// TIA Portal V21 export
// export: Created 2026-10-23T20:42:47.6019008Z, ExportSetting WithDefaults, DisplayName Totally Integrated Automation Portal, DisplayVersion V21 Update 1, DisplayName SINAMICS Startdrive Advanced, DisplayVersion V21 HF2, DisplayName SINAMICS Startdrive G110M, G120, G120C, G120D, G120P, G115D, DisplayVersion V21 HF2, DisplayName SINAMICS Startdrive G130, G150, S120, S150, G200, G220, S200, S210, S220, Innomotics MVD, DisplayVersion V21 HF2, DisplayName STEP 7 Professional, DisplayVersion V21 Update 1, DisplayName STEP 7 Safety, DisplayVersion V21, DisplayName Tech WebApplication, DisplayVersion V21, DisplayName WinCC Basic/Comfort/Advanced, DisplayVersion V21 Update 1, DisplayName WinCC Unified, DisplayVersion V21 Update 1
FUNCTION_BLOCK "FB_FbdBoxes"   // FB10, FBD
TITLE = FUP-Boxen, Aufruf und Sprung / FBD boxes, call and jump
{ S7_Optimized_Access := 'TRUE' }
VERSION : 0.1
// TON, MOVE, ADD, Vergleich, FB-Aufruf mit EN/ENO und ein Sprung mit Marke in FUP / TON, MOVE, ADD, compare, FB call with EN/ENO and a jump with label in FBD
// stored: AutoNumber true, IsIECCheckEnabled false, IsRetainMemResEnabled false, MemoryReserve 100, SetENOAutomatically false, UDAEnableTagReadback false
   VAR_INPUT
      Start : Bool;   // Startbefehl / Start command
      InValue : Int;   // Eingangswert / Input value
      Limit : Int := 100;   // Grenzwert für den Vergleich / Limit for the comparison
   END_VAR
   VAR_OUTPUT
      Delayed : Bool;   // Start um drei Sekunden verzögert / Start delayed by three seconds
      Copy : Int;   // Kopie des Eingangswerts / Copy of the input value
      Sum : Int;   // Eingangswert plus Grenzwert / Input value plus limit
      IsEqual : Bool;   // Eingangswert gleich dem Grenzwert / Input value equal to the limit
      SectionsOk : Bool;   // ENO des Aufrufs von FB_SclTimers / ENO of the FB_SclTimers call
      Skipped : Bool;   // Nur gesetzt, wenn nicht gesprungen wird / Set only when the jump is not taken
      AfterJump : Bool;   // Netzwerk nach der Sprungmarke / Network after the jump label
   END_VAR
   VAR
      Delay { S7_SetPoint := 'True'} : TON_TIME;   // Einschaltverzögerung / On-delay timer
      DelayElapsed : Time;   // Abgelaufene Zeit der Einschaltverzögerung / Elapsed time of the on-delay timer
      Timers { S7_SetPoint := 'True'} : "FB_SclTimers";   // Multiinstanz von FB_SclTimers / Multi-instance of FB_SclTimers
      TimerRunOn : Bool;   // Nachlaufausgang von FB_SclTimers / Run-on output of FB_SclTimers
      TimerPulse : Bool;   // Impulsausgang von FB_SclTimers / Pulse output of FB_SclTimers
      TimerCount : Int;   // Zählausgang von FB_SclTimers / Count output of FB_SclTimers
      TimerDelayed : Bool;   // Verzögerter Ausgang von FB_SclTimers / Delayed output of FB_SclTimers
      TimerReached : Bool;   // Ausgang Zählwert erreicht von FB_SclTimers / Count reached output of FB_SclTimers
   END_VAR
   VAR_TEMP   // added for the SCL form of the ladder/FBD networks
      _w1 : Bool;
   END_VAR
BEGIN

REGION Network 1: Einschaltverzögerung als Multiinstanz / On-delay timer as multi-instance
   // Der Ausgang folgt dem Startbefehl nach drei Sekunden. / The output follows the start command after three seconds.
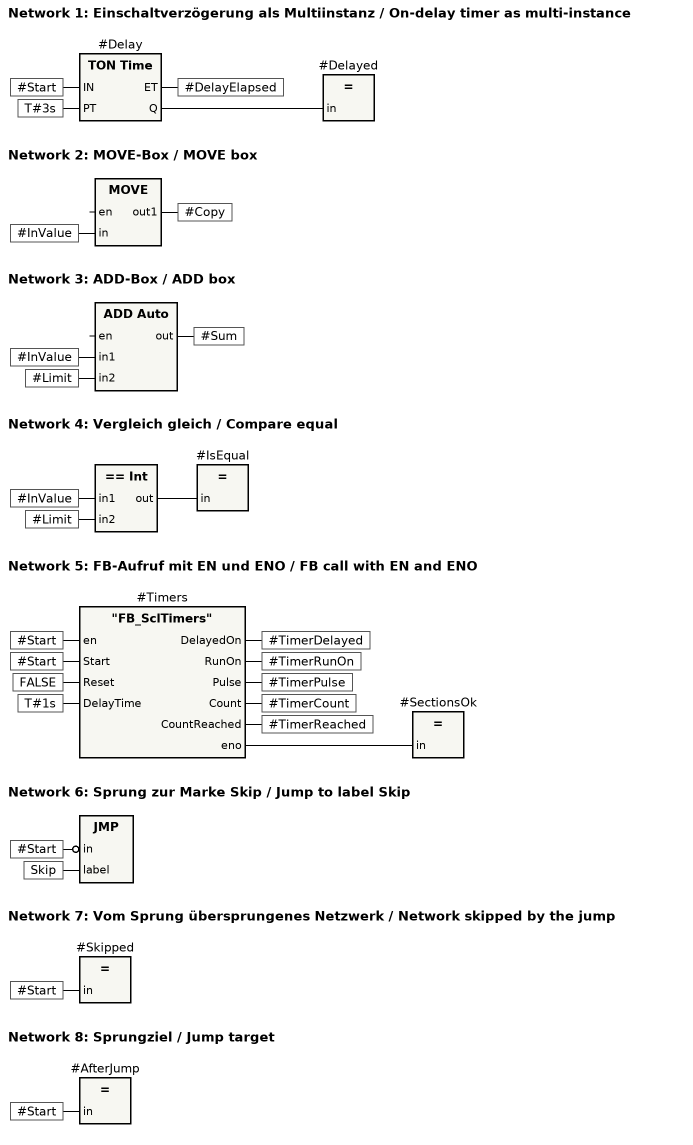
   #Delay(IN := #Start, PT := T#3s, ET => #DelayElapsed);   // TON
   #Delayed := #Delay.Q;
END_REGION

REGION Network 2: MOVE-Box / MOVE box
   // Kopiert den Eingangswert. / Copies the input value.
   #Copy := #InValue;
END_REGION

REGION Network 3: ADD-Box / ADD box
   // Addiert den Grenzwert zum Eingangswert. / Adds the limit to the input value.
   #Sum := #InValue + #Limit;
END_REGION

REGION Network 4: Vergleich gleich / Compare equal
   // Wahr, wenn der Eingangswert dem Grenzwert entspricht. / True when the input value equals the limit.
   #IsEqual := #InValue = #Limit;
END_REGION

REGION Network 5: FB-Aufruf mit EN und ENO / FB call with EN and ENO
   // Ruft FB_SclTimers als Multiinstanz auf, wenn Start an ist. / Calls FB_SclTimers as a multi-instance when start is on.
   #Timers(EN := #Start,   // "FB_SclTimers"
           Start := #Start,
           Reset := FALSE,
           DelayTime := T#1s,
           DelayedOn => #TimerDelayed,
           RunOn => #TimerRunOn,
           Pulse => #TimerPulse,
           Count => #TimerCount,
           CountReached => #TimerReached,
           ENO => #_w1);
   #SectionsOk := #_w1;
END_REGION

REGION Network 6: Sprung zur Marke Skip / Jump to label Skip
   // Springt über das nächste Netzwerk, wenn Start aus ist. / Jumps over the next network when start is off.
   IF NOT #Start THEN GOTO Skip; END_IF;
END_REGION

REGION Network 7: Vom Sprung übersprungenes Netzwerk / Network skipped by the jump
   // Läuft nur, wenn nicht gesprungen wird. / Runs only when the jump is not taken.
   #Skipped := #Start;
END_REGION

REGION Network 8: Sprungziel / Jump target
   // Die Marke Skip kennzeichnet dieses Netzwerk. / The label Skip marks this network.
   Skip:
   #AfterJump := #Start;
END_REGION
END_FUNCTION_BLOCK
